// TIA Portal V21 export
// export: Created 2026-10-23T20:42:56.9111518Z, ExportSetting WithDefaults, DisplayName Totally Integrated Automation Portal, DisplayVersion V21 Update 1, DisplayName SINAMICS Startdrive Advanced, DisplayVersion V21 HF2, DisplayName SINAMICS Startdrive G110M, G120, G120C, G120D, G120P, G115D, DisplayVersion V21 HF2, DisplayName SINAMICS Startdrive G130, G150, S120, S150, G200, G220, S200, S210, S220, Innomotics MVD, DisplayVersion V21 HF2, DisplayName STEP 7 Professional, DisplayVersion V21 Update 1, DisplayName STEP 7 Safety, DisplayVersion V21, DisplayName Tech WebApplication, DisplayVersion V21, DisplayName WinCC Basic/Comfort/Advanced, DisplayVersion V21 Update 1, DisplayName WinCC Unified, DisplayVersion V21 Update 1
DATA_BLOCK "DB_CallData"   // DB17
TITLE = Call data of OB_Main
{ S7_Optimized_Access := 'TRUE' }
VERSION : 0.1
// Actual parameters of the FC calls in OB_Main that must persist between cycles
// stored: AutoNumber true, DBAccessibleFromOPCUA true, DBAccessibleFromWebserver true, IsOnlyStoredInLoadMemory false, IsRetainMemResEnabled false, IsWriteProtectedInAS false, MemoryReserve 100
   VAR
      Values : Array[0..9] of Real;   // Values for FB_SclCalls
      LadMotor : Bool;   // Output Motor of FC_LadContacts
      LadPulse : Bool;   // Output Pulse of FC_LadContacts
      LadFallingPulse : Bool;   // Output FallingPulse of FC_LadContacts
      LadAlarm : Bool;   // Output Alarm of FC_LadContacts
      LadLamp : Bool;   // Output Lamp of FC_LadContacts
      LadBranch : Bool;   // Output BranchResult of FC_LadContacts
      LadLatched : Bool;   // InOut Latched of FC_LadContacts
      LadRiseMemory : Bool;   // Edge memory for FC_LadContacts
      LadFallMemory : Bool;   // Edge memory for FC_LadContacts
      LadCoilMemory : Bool;   // Edge memory for FC_LadContacts
      FbdAnd : Bool;   // Output AndOut of FC_FbdLogic
      FbdOr : Bool;   // Output OrOut of FC_FbdLogic
      FbdXor : Bool;   // Output XorOut of FC_FbdLogic
      FbdNot : Bool;   // Output NotOut of FC_FbdLogic
      FbdSr : Bool;   // Output SrOut of FC_FbdLogic
      FbdRs : Bool;   // Output RsOut of FC_FbdLogic
      FbdEdge : Bool;   // Output EdgeOut of FC_FbdLogic
      FbdSrBit : Bool;   // InOut SrBit of FC_FbdLogic
      FbdRsBit : Bool;   // InOut RsBit of FC_FbdLogic
      FbdEdgeBit : Bool;   // InOut EdgeBit of FC_FbdLogic
   END_VAR
BEGIN
END_DATA_BLOCK
